{attribute 'qualified_only'}
{attribute 'strict'}
TYPE E_Stirrer_mode :
(
	off := 0,
	continues,
	cyclic
);
END_TYPE

(* stored: Version 1.1.0.1, ProductVersion 3.1.4024.13
   DUT E_Stirrer_mode: Id {1da0c747-f172-416a-940f-6936dbbbb95c} *)
